// TIA Portal V15.1 export
// export: Created 2026-09-17T17:40:09.8316095Z, ExportSetting WithDefaults, DisplayName Totally Integrated Automation Portal, DisplayVersion V15.1, DisplayName TIA Portal Openness, DisplayVersion V15.1, DisplayName STEP 7 Professional, DisplayVersion V15.1, DisplayName WinCC Professional, DisplayVersion V15.1
Screen "Start Screen"  1024x768, Number=1
  ScreenLayer 
    GraphicView "Graphic view_1" at 0,1 size 1016x767  Picture=images (5)
    GraphicView "Graphic view_2" at 818,8 size 158x89  Picture=Graphic_1
    TextField "Text field_1" at 793,97 size 231x21  Text="By Ahmad Saber Zain"
    Button "Button_1" at 31,675 size 90x44  Mode=Text, StyleItem=Button, TextOff="End RT", TextOn="Text"
      on Press: StopRuntime(Mode := 0)
    Button "Button_2" at 31,619 size 90x44  Mode=Text, StyleItem=Button, TextOff="Trolley", TextOn="Text"
      on Press: ActivateScreen(Screen name := Trolley, Object number := 0)
    Button "Button_3" at 31,565 size 90x44  Mode=Text, StyleItem=Button, TextOff="Slewing", TextOn="Text"
      on Press: ActivateScreen(Screen name := slewing, Object number := 0)
    Button "Button_4" at 31,511 size 90x44  Mode=Text, StyleItem=Button, TextOff="Hook", TextOn="Text"
      on Press: ActivateScreen(Screen name := Hook, Object number := 0)
    Button "Button_5" at 31,457 size 90x44  Mode=Text, StyleItem=Button, TextOff="Faults", TextOn="Text"
      on Press: ActivateScreen(Screen name := faults, Object number := 0)
    Button "Button_6" at 31,403 size 90x44  Mode=Text, StyleItem=Button, TextOff="Motion", TextOn="Text"
      on Press: ActivateScreen(Screen name := Motion, Object number := 0)
    TextField "Text field_2" at 618,8 size 163x29  Text="Start Screen"
